Fanuc KAREL source: kd00044.KL

PROGRAM KD00044
%STACKSIZE=65535
%PRIORITY=65535
%NOLOCKGROUP
VAR
I : INTEGER
J : INTEGER
B : BOOLEAN
R : REAL
S : STRING[80]
-- UNRESOLVED DECLARATIONS (source type spelling not recovered)
-- G : TYPE_0x011E (type_u16=0x011E)
BEGIN
I=1
END KD00044
